(* IEC 61131-3 sources: codesys-to-astra/src/POUs/F_C2aAddChar, 2 files *)

(* ---- F_C2aAddChar.decl.st ---- *)
// Назначение: замена OSU.ADD_CHAR (OwenStringUtils v3.0, с. 33): дополнение sInputString символом sAddChar
//             до длины usiTargetLen справа (xRight) или слева; длиннее — без изменений.
// Автор:      kr0nsch
// Версия:     0.1.0
// Документ:   docs/LIBMAP.md
FUNCTION F_C2aAddChar : STRING(255)
VAR_INPUT
    sInputString : STRING(255); // исходная строка
    usiTargetLen : USINT;       // длина результата
    sAddChar : STRING(1);       // символ-заполнитель
    xRight : BOOL;              // TRUE — справа, FALSE — слева
END_VAR
VAR
    sResult : STRING(255);  // результат
    iGuard : INT;           // защита от бесконечного цикла при пустом sAddChar
END_VAR

(* ---- F_C2aAddChar.impl.st ---- *)
sResult := sInputString;
iGuard := 0;
WHILE LEN(sResult) < USINT_TO_INT(usiTargetLen) AND LEN(sAddChar) > 0
        AND iGuard < 255 DO  // lint:allow STL008 STRING(255)
    IF xRight THEN
        sResult := CONCAT(sResult, sAddChar);
    ELSE
        sResult := CONCAT(sAddChar, sResult);
    END_IF
    iGuard := iGuard + 1;
END_WHILE
F_C2aAddChar := sResult;
